FUNCTION_BLOCK DUTY_STANDBY (* Migrated from IEC 61131-3 ST *)
  (* Standard: 61499-2 *)
  (* Version 1.0, 2026-11-06, st2fb *)
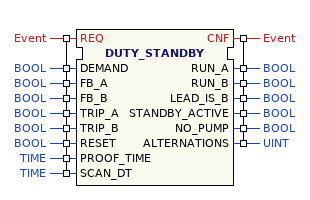
  EVENT_INPUT
    REQ WITH DEMAND, FB_A, FB_B, TRIP_A, TRIP_B, RESET, PROOF_TIME, SCAN_DT;
  END_EVENT
  EVENT_OUTPUT
    CNF WITH RUN_A, RUN_B, LEAD_IS_B, STANDBY_ACTIVE, NO_PUMP, ALTERNATIONS;
  END_EVENT
  VAR_INPUT
    DEMAND : BOOL;
    FB_A : BOOL;
    FB_B : BOOL;
    TRIP_A : BOOL;
    TRIP_B : BOOL;
    RESET : BOOL;
    PROOF_TIME : TIME;
    SCAN_DT : TIME;
  END_VAR
  VAR_OUTPUT
    RUN_A : BOOL;
    RUN_B : BOOL;
    LEAD_IS_B : BOOL;
    STANDBY_ACTIVE : BOOL;
    NO_PUMP : BOOL;
    ALTERNATIONS : UINT;
  END_VAR
  VAR
    ST2FB_NOW : TIME := T#0s;
    DEMAND_END_CLK : BOOL;
    DEMAND_END_Q : BOOL;
    DEMAND_END_M : BOOL;
    PROOF_A_IN : BOOL;
    PROOF_A_PT : TIME;
    PROOF_A_Q : BOOL;
    PROOF_A_ET : TIME;
    PROOF_A_STATE : INT;
    PROOF_A_PREV_IN : BOOL;
    PROOF_A_START_TIME : TIME;
    PROOF_B_IN : BOOL;
    PROOF_B_PT : TIME;
    PROOF_B_Q : BOOL;
    PROOF_B_ET : TIME;
    PROOF_B_STATE : INT;
    PROOF_B_PREV_IN : BOOL;
    PROOF_B_START_TIME : TIME;
    FAILED_A_S1 : BOOL;
    FAILED_A_R : BOOL;
    FAILED_A_Q1 : BOOL;
    FAILED_B_S1 : BOOL;
    FAILED_B_R : BOOL;
    FAILED_B_Q1 : BOOL;
  END_VAR
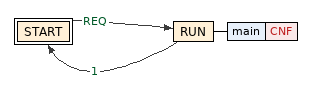
  EC_STATES
    START;
    RUN : main -> CNF;
  END_STATES
  EC_TRANSITIONS
    START TO RUN := REQ;
    RUN TO START := 1;
  END_TRANSITIONS
  ALGORITHM main IN ST:
ST2FB_NOW := ST2FB_NOW + SCAN_DT;

DEMAND_END_CLK := DEMAND;
DEMAND_END_Q := NOT DEMAND_END_CLK AND NOT DEMAND_END_M;
DEMAND_END_M := NOT DEMAND_END_CLK;
IF DEMAND_END_Q THEN
  LEAD_IS_B := NOT LEAD_IS_B;
  ALTERNATIONS := ALTERNATIONS + 1;
END_IF;

PROOF_A_IN := RUN_A AND NOT FB_A;
PROOF_A_PT := PROOF_TIME;
IF (PROOF_A_STATE = 0) AND NOT PROOF_A_PREV_IN AND PROOF_A_IN THEN
  PROOF_A_STATE := 1;
  PROOF_A_Q := FALSE;
  PROOF_A_START_TIME := ST2FB_NOW;
ELSE
  IF NOT PROOF_A_IN THEN
    PROOF_A_ET := T#0s;
    PROOF_A_Q := FALSE;
    PROOF_A_STATE := 0;
  ELSIF PROOF_A_STATE = 1 THEN
    IF PROOF_A_START_TIME + PROOF_A_PT <= ST2FB_NOW THEN
      PROOF_A_STATE := 2;
      PROOF_A_Q := TRUE;
      PROOF_A_ET := PROOF_A_PT;
    ELSE
      PROOF_A_ET := ST2FB_NOW - PROOF_A_START_TIME;
    END_IF;
  END_IF;
END_IF;
PROOF_A_PREV_IN := PROOF_A_IN;

PROOF_B_IN := RUN_B AND NOT FB_B;
PROOF_B_PT := PROOF_TIME;
IF (PROOF_B_STATE = 0) AND NOT PROOF_B_PREV_IN AND PROOF_B_IN THEN
  PROOF_B_STATE := 1;
  PROOF_B_Q := FALSE;
  PROOF_B_START_TIME := ST2FB_NOW;
ELSE
  IF NOT PROOF_B_IN THEN
    PROOF_B_ET := T#0s;
    PROOF_B_Q := FALSE;
    PROOF_B_STATE := 0;
  ELSIF PROOF_B_STATE = 1 THEN
    IF PROOF_B_START_TIME + PROOF_B_PT <= ST2FB_NOW THEN
      PROOF_B_STATE := 2;
      PROOF_B_Q := TRUE;
      PROOF_B_ET := PROOF_B_PT;
    ELSE
      PROOF_B_ET := ST2FB_NOW - PROOF_B_START_TIME;
    END_IF;
  END_IF;
END_IF;
PROOF_B_PREV_IN := PROOF_B_IN;

FAILED_A_S1 := TRIP_A OR PROOF_A_Q;
FAILED_A_R := RESET;
FAILED_A_Q1 := FAILED_A_S1 OR (NOT FAILED_A_R AND FAILED_A_Q1);

FAILED_B_S1 := TRIP_B OR PROOF_B_Q;
FAILED_B_R := RESET;
FAILED_B_Q1 := FAILED_B_S1 OR (NOT FAILED_B_R AND FAILED_B_Q1);

RUN_A := DEMAND AND NOT FAILED_A_Q1 AND (NOT LEAD_IS_B OR FAILED_B_Q1);
RUN_B := DEMAND AND NOT FAILED_B_Q1 AND (LEAD_IS_B OR FAILED_A_Q1);
STANDBY_ACTIVE := (RUN_A AND LEAD_IS_B) OR (RUN_B AND NOT LEAD_IS_B);
NO_PUMP := DEMAND AND FAILED_A_Q1 AND FAILED_B_Q1;
  END_ALGORITHM
END_FUNCTION_BLOCK
